TEXTLIST TextList_Piston_Recipe_State_OpenClose
  0 = ' '
  1 = 'Open'
  2 = 'Close'
   = ''
END_TEXTLIST

(* stored: Version 1.1.0.1, ProductVersion 3.1.4024.12
   TextList TextList_Piston_Recipe_State_OpenClose: Id {999aad2f-a4fd-427b-be34-9b9abe26f1b3} *)
